// TIA Portal V20 export
// export: Created 2026-10-20T18:55:47.0251742Z, ExportSetting None, DisplayName Totally Integrated Automation Portal, DisplayVersion V20 Update 6, DisplayName TIA Portal Openness, DisplayVersion V20 Update 6, DisplayName TIA Portal Version Control Interface, DisplayVersion V20 Update 6, DisplayName SINAMICS Startdrive Advanced, DisplayVersion V20 SP1, DisplayName SINAMICS Startdrive G130, G150, S120, S150, SINAMICS MV, G220, S200, S210, DisplayVersion V20 SP1, DisplayName SINAMICS Startdrive G110M, G120, G120C, G120D, G120P, G115D, DisplayVersion V20 SP1, DisplayName STEP 7 Professional, DisplayVersion V20 Update 6, DisplayName STEP 7 Safety, DisplayVersion V20 Update 2, DisplayName WinCC Basic/Comfort/Advanced, DisplayVersion V20 Update 6, DisplayName WinCC Unified, DisplayVersion V20 Update 6
VAR_GLOBAL   // PLC tag table "Lock_4"
   "Lock Reset_4" AT %Q1362.0 : Bool;
   Switches_4 AT %IB1164 : Byte;
   Lock_4_Estop_CH2 AT %I1782.3 : Bool;
   Lamps_4 AT %QB1079 : Byte;
   Lock_4_Closed_CH2 AT %I1782.1 : Bool;
   Lock_4_Estop_CH1 AT %I1782.2 : Bool;
   Lock_4_Closed_CH1 AT %I1782.0 : Bool;
   "Solenoid Enable_4" AT %Q1080.0 : Bool;
   Lock_4_Reset_Input3 AT %Q1783.2 : Bool;
   Lock_4_Reset_Input4 AT %Q1783.3 : Bool;
   Lock_4_Reset_Input2 AT %Q1783.1 : Bool;
   Lock_4_Reset_Input1 AT %Q1783.0 : Bool;
   "Guard Position_4" AT %I1199.0 : Bool;
   "Lock Position_4" AT %I1200.0 : Bool;
END_VAR
